(* IEC 61131-3 sources: kns-port-domestic/targets/astra/lib/src/DUTs/Valve, 7 files *)

(* ---- E_ValveAlarm.dut.st ---- *)
// Назначение: индексы слотов тревог запорной арматуры. Нестрогое перечисление: им
//             индексируются массивы.
// Автор:      kr0nsch
// Версия:     0.1.0
// Документ:   docs/fb/FB_Valve.md
{attribute 'qualified_only'}
TYPE E_ValveAlarm :
(
    FailToOpen   := 0,   // не открылась за tTravel
    FailToClose  := 1,   // не закрылась за tTravel
    BothLimits   := 2,   // оба концевика
    PositionLost := 3,   // уход с концевика без команды
    TorqueTrip   := 4,   // муфта в ходе
    ExtFault     := 5,   // авария привода
    InterlockAct := 6    // действует блокировка (по умолчанию выключена)
) UINT;
END_TYPE

(* ---- E_ValveSafePos.dut.st ---- *)
// Назначение: куда вести арматуру по защитной блокировке.
// Автор:      kr0nsch
// Версия:     0.1.0
// Документ:   docs/fb/FB_Valve.md
{attribute 'qualified_only'}
{attribute 'strict'}
TYPE E_ValveSafePos :
(
    Closed := 0,   // закрыть
    Open   := 1,   // открыть
    Stay   := 2    // остановить (только Motorized)
) INT;
END_TYPE

(* ---- E_ValveState.dut.st ---- *)
// Назначение: состояние запорной арматуры.
// Автор:      kr0nsch
// Версия:     0.1.0
// Документ:   docs/fb/FB_Valve.md
{attribute 'qualified_only'}
{attribute 'strict'}
TYPE E_ValveState :
(
    Unknown      := 0,   // нет концевиков и нет истории
    Closed       := 1,
    Opening      := 2,
    Open         := 3,
    Closing      := 4,
    Intermediate := 5,   // остановлена в промежутке
    Reversing    := 6,   // пауза перед сменой направления
    Fault        := 7
) INT;
END_TYPE

(* ---- E_ValveType.dut.st ---- *)
// Назначение: вид запорной арматуры: соленоид с пружинным возвратом или электропривод.
// Автор:      kr0nsch
// Версия:     0.1.0
// Документ:   docs/fb/FB_Valve.md
{attribute 'qualified_only'}
{attribute 'strict'}
TYPE E_ValveType :
(
    SolenoidEto := 0,   // соленоид, «под током — открыт» (НЗ клапан); без тока — закрыт
    SolenoidEtc := 1,   // соленоид, «под током — закрыт» (НО клапан); без тока — открыт
    Motorized   := 2    // электропривод: выходы «открывать»/«закрывать», стоп в промежутке
) INT;
END_TYPE

(* ---- ST_ValveCfg.dut.st ---- *)
// Назначение: параметры запорной арматуры (Persistent Variables приложения,
//             VAR_IN_OUT CONSTANT stCfg). Значения по умолчанию проходят CheckConfig.
//             Тип лежит в Persistent Variables приложения и заморожен в пределах 1.x (A-13).
// Автор:      kr0nsch
// Версия:     0.1.0
// Документ:   docs/fb/FB_Valve.md
{attribute 'qualified_only'}
TYPE ST_ValveCfg :
STRUCT
    eType            : E_ValveType := E_ValveType.Motorized;
    xZsoUsed         : BOOL := TRUE;      // концевик «открыто» подключён
    xZscUsed         : BOOL := TRUE;      // концевик «закрыто» подключён
    tTravel          : TIME := T#60S;     // макс. время хода (паспорт привода + запас); без концевика — «по времени»
    tLimitFilter     : TIME := T#500MS;   // фильтр «оба концевика» и ухода с концевика
    tReverse         : TIME := T#1S;      // пауза перед реверсом (Motorized)
    xTorqueUsed      : BOOL := FALSE;     // муфта подключена (Motorized)
    xCloseOnTorque   : BOOL := FALSE;     // закрытие «по моменту» (клиновые задвижки)
    eSafePos         : E_ValveSafePos := E_ValveSafePos.Closed;   // куда вести по блокировке
    wInterlockMask   : WORD := 16#FFFF;   // какие биты wInterlock действуют
    wPermitOpenMask  : WORD := 16#FFFF;   // какие биты wPermitOpen обязательны для открытия
    wPermitCloseMask : WORD := 16#FFFF;   // какие биты wPermitClose обязательны для закрытия
    tResetWindow     : TIME := T#3S;      // окно снятия причин после Reset
    udiMaintCycles   : UDINT := 0;        // ТО по числу циклов; 0 — нет
    udiAlarmIdBase   : UDINT := 0;        // номер первой тревоги устройства (dev_no * 10)
    astAlarm         : ARRAY[0..GVL_Const.DEV_ALARMS_MAX - 1] OF ST_AlarmCfg := [
        (ePriority := E_AlarmPriority.Medium),    // 0 FailToOpen
        (ePriority := E_AlarmPriority.Medium),    // 1 FailToClose
        (ePriority := E_AlarmPriority.Medium),    // 2 BothLimits
        (ePriority := E_AlarmPriority.Medium),    // 3 PositionLost
        (ePriority := E_AlarmPriority.Medium),    // 4 TorqueTrip
        (ePriority := E_AlarmPriority.Medium),    // 5 ExtFault
        (ePriority := E_AlarmPriority.None),      // 6 InterlockAct
        (ePriority := E_AlarmPriority.None)];     // 7 —
END_STRUCT
END_TYPE

(* ---- ST_ValveCmd.dut.st ---- *)
// Назначение: команды HMI/SCADA запорной арматуры (GVL_Hmi приложения, VAR_IN_OUT stCmd).
// Автор:      kr0nsch
// Версия:     0.1.0
// Документ:   docs/fb/FB_Valve.md
{attribute 'qualified_only'}
TYPE ST_ValveCmd :
STRUCT
    stCommon    : ST_DeviceCmd;
    xOpen       : BOOL;   // импульс: открыть (в Auto — переход в Manual и открыть)
    xClose      : BOOL;   // импульс: закрыть (в Auto — переход в Manual и закрыть)
    xStop       : BOOL;   // импульс: стоп (только Motorized; в Auto — переход в Manual)
    xResetMaint : BOOL;   // импульс: обнулить счётчики «с последнего ТО»
END_STRUCT
END_TYPE

(* ---- ST_ValveSts.dut.st ---- *)
// Назначение: состояние запорной арматуры для HMI/SCADA. 52 байта, 26 регистров Modbus:
//             только 16- и 32-битные поля без скрытого выравнивания.
// Автор:      kr0nsch
// Версия:     0.1.0
// Документ:   docs/fb/FB_Valve.md
{attribute 'qualified_only'}
TYPE ST_ValveSts :
STRUCT
    stCommon         : ST_DeviceSts;   // 0..27
    eState           : E_ValveState;   // 28
    wInterlock       : WORD;     // 30: действующие блокировки (после маски)
    wPermitMissing   : WORD;     // 32: недостающие разрешения для текущего направления
    uiFirstOut       : UINT;     // 34: первопричина блокировки; NO_FIRST_OUT — нет
    uiTravelRemain_s : UINT;     // 36: до таймаута хода, с
    wReserve         : WORD;     // 38: выравнивание следующего 32-битного поля
    udiCycles        : UDINT;    // 40: циклов «открыто» всего
    udiCyclesMaint   : UDINT;    // 44: с последнего ТО
    rActTime_h       : REAL;     // 48: время работы привода, ч
END_STRUCT
END_TYPE
